(* IEC 61131-3 sources: plc-iiot-stack/tests/DUTs, 2 files *)

(* ---- ST_FakeMqttIn.dut.st ---- *)
// Назначение: входящее сообщение в очереди подменного клиента FB_MqttClientFake.
// Документ:   docs/TEST_REPORT.md
{attribute 'qualified_only'}
TYPE ST_FakeMqttIn :
STRUCT
    sTopic : STRING(GVL_Const.MQTT_TOPIC_LEN);
    sPayload : STRING(GVL_Const.MQTT_CMD_PAYLOAD_LEN);
    xTruncated : BOOL;
    xRetained : BOOL;
END_STRUCT
END_TYPE

(* ---- ST_FakeMqttMsg.dut.st ---- *)
// Назначение: сообщение, опубликованное через подменный клиент FB_MqttClientFake.
// Документ:   docs/TEST_REPORT.md
{attribute 'qualified_only'}
TYPE ST_FakeMqttMsg :
STRUCT
    sTopic : STRING(GVL_Const.MQTT_TOPIC_LEN);
    sPayload : STRING(GVL_Const.MQTT_PAYLOAD_LEN);
    eQos : E_MqttQos;
    xRetain : BOOL;
END_STRUCT
END_TYPE
